// TIA Portal V20 export
// export: Created 2026-10-12T16:46:21.2512709Z, ExportSetting WithDefaults, DisplayName Totally Integrated Automation Portal, DisplayVersion V20 Update 6, DisplayName TIA Portal Openness, DisplayVersion V20 Update 6, DisplayName TIA Portal Version Control Interface, DisplayVersion V20 Update 6, DisplayName SINAMICS Startdrive Advanced, DisplayVersion V20 SP1 Update 2, DisplayName SINAMICS Startdrive G110M, G120, G120C, G120D, G120P, G115D, DisplayVersion V20 SP1 Update 2, DisplayName SINAMICS Startdrive G130, G150, S120, S150, SINAMICS MV, G220, S200, S210, DisplayVersion V20 SP1 Update 2, DisplayName STEP 7 Professional, DisplayVersion V20 Update 6, DisplayName STEP 7 Safety, DisplayVersion V20 Update 2, DisplayName WinCC Basic/Comfort/Advanced, DisplayVersion V20 Update 6, DisplayName WinCC Professional, DisplayVersion V20 Update 6, DisplayName WinCC Unified, DisplayVersion V20 Update 6
ORGANIZATION_BLOCK "Main"   // OB1, LAD, ProgramCycle
TITLE = "Main Program Sweep (Cycle)"
{ S7_Optimized_Access := 'TRUE' }
VERSION : 0.1
// stored: AutoNumber true, IsIECCheckEnabled false, SetENOAutomatically false
   VAR_INPUT
      Initial_Call : Bool;   // Initial call of this OB
      Remanence : Bool;   // =True, if remanent data are available
   END_VAR
   VAR_TEMP
      Lampentest_Ein : Bool;
      Blinktakt : Bool;
   END_VAR
BEGIN

REGION Network 1 (SCL): Eingaenge Lesen
   //KP8_1
   "FB_KP8_DB_1".KP8.Rohdaten.IB_Tasten := "KP8_1_IB_Tasten";
   "FB_KP8_DB_1".KP8.Rohdaten.IB_DI := "KP8_1_IB_DI";
   "FB_KP8_DB_1"();

   //KP8_2
   "FB_KP8_DB_2".KP8.Rohdaten.IB_Tasten := "KP8_2_IB_Tasten";
   "FB_KP8_DB_2".KP8.Rohdaten.IB_DI := "KP8_2_IB_DI";
   "FB_KP8_DB_2"();

   //KP8_3
   "FB_KP8_DB_3".KP8.Rohdaten.IB_Tasten := "KP8_3_IB_Tasten";
   "FB_KP8_DB_3".KP8.Rohdaten.IB_DI := "KP8_3_IB_DI";
   "FB_KP8_DB_3"();

   //KP8_4
   "FB_KP8_DB_4".KP8.Rohdaten.IB_Tasten := "KP8_4_IB_Tasten";
   "FB_KP8_DB_4".KP8.Rohdaten.IB_DI := "KP8_4_IB_DI";
   "FB_KP8_DB_4"();

   //KP8_5
   "FB_KP8_DB_5".KP8.Rohdaten.IB_Tasten := "KP8_5_IB_Tasten";
   "FB_KP8_DB_5".KP8.Rohdaten.IB_DI := "KP8_5_IB_DI";
   "FB_KP8_DB_5"();

   //KP8_6
   "FB_KP8_DB_6".KP8.Rohdaten.IB_Tasten := "KP8_6_IB_Tasten";
   "FB_KP8_DB_6".KP8.Rohdaten.IB_DI := "KP8_6_IB_DI";
   "FB_KP8_DB_6"();

   //KP8_7
   "FB_KP8_DB_7".KP8.Rohdaten.IB_Tasten := "KP8_7_IB_Tasten";
   "FB_KP8_DB_7".KP8.Rohdaten.IB_DI := "KP8_7_IB_DI";
   "FB_KP8_DB_7"();

   //KP8_8
   "FB_KP8_DB_8".KP8.Rohdaten.IB_Tasten := "KP8_8_IB_Tasten";
   "FB_KP8_DB_8".KP8.Rohdaten.IB_DI := "KP8_8_IB_DI";
   "FB_KP8_DB_8"();

   //KP8_9
   "FB_KP8_DB_9".KP8.Rohdaten.IB_Tasten := "KP8_9_IB_Tasten";
   "FB_KP8_DB_9".KP8.Rohdaten.IB_DI := "KP8_9_IB_DI";
   "FB_KP8_DB_9"();

   //KP8_10
   "FB_KP8_DB_10".KP8.Rohdaten.IB_Tasten := "KP8_10_IB_Tasten";
   "FB_KP8_DB_10".KP8.Rohdaten.IB_DI := "KP8_10_IB_DI";
   "FB_KP8_DB_10"();

   //KP8_11
   "FB_KP8_DB_11".KP8.Rohdaten.IB_Tasten := "KP8_11_IB_Tasten";
   "FB_KP8_DB_11".KP8.Rohdaten.IB_DI := "KP8_11_IB_DI";
   "FB_KP8_DB_11"();

   //KP8_12
   "FB_KP8_DB_12".KP8.Rohdaten.IB_Tasten := "KP8_12_IB_Tasten";
   "FB_KP8_DB_12".KP8.Rohdaten.IB_DI := "KP8_12_IB_DI";
   "FB_KP8_DB_12"();

   //KP8_13
   "FB_KP8_DB_13".KP8.Rohdaten.IB_Tasten := "KP8_13_IB_Tasten";
   "FB_KP8_DB_13".KP8.Rohdaten.IB_DI := "KP8_13_IB_DI";
   "FB_KP8_DB_13"();

   //KP8_14
   "FB_KP8_DB_14".KP8.Rohdaten.IB_Tasten := "KP8_14_IB_Tasten";
   "FB_KP8_DB_14".KP8.Rohdaten.IB_DI := "KP8_14_IB_DI";
   "FB_KP8_DB_14"();

   //KP8_15
   "FB_KP8_DB_15".KP8.Rohdaten.IB_Tasten := "KP8_15_IB_Tasten";
   "FB_KP8_DB_15".KP8.Rohdaten.IB_DI := "KP8_15_IB_DI";
   "FB_KP8_DB_15"();

   //KP8_16
   "FB_KP8_DB_16".KP8.Rohdaten.IB_Tasten := "KP8_16_IB_Tasten";
   "FB_KP8_DB_16".KP8.Rohdaten.IB_DI := "KP8_16_IB_DI";
   "FB_KP8_DB_16"();

   //KP8_17
   "FB_KP8_DB_17".KP8.Rohdaten.IB_Tasten := "KP8_17_IB_Tasten";
   "FB_KP8_DB_17".KP8.Rohdaten.IB_DI := "KP8_17_IB_DI";
   "FB_KP8_DB_17"();

   //KP8_18
   "FB_KP8_DB_18".KP8.Rohdaten.IB_Tasten := "KP8_18_IB_Tasten";
   "FB_KP8_DB_18".KP8.Rohdaten.IB_DI := "KP8_18_IB_DI";
   "FB_KP8_DB_18"();

   //KP8_19
   "FB_KP8_DB_19".KP8.Rohdaten.IB_Tasten := "KP8_19_IB_Tasten";
   "FB_KP8_DB_19".KP8.Rohdaten.IB_DI := "KP8_19_IB_DI";
   "FB_KP8_DB_19"();

   //KP8_20
   "FB_KP8_DB_20".KP8.Rohdaten.IB_Tasten := "KP8_20_IB_Tasten";
   "FB_KP8_DB_20".KP8.Rohdaten.IB_DI := "KP8_20_IB_DI";
   "FB_KP8_DB_20"();

   //KP8_21
   "FB_KP8_DB_21".KP8.Rohdaten.IB_Tasten := "KP8_21_IB_Tasten";
   "FB_KP8_DB_21".KP8.Rohdaten.IB_DI := "KP8_21_IB_DI";
   "FB_KP8_DB_21"();

   //KP8_22
   "FB_KP8_DB_22".KP8.Rohdaten.IB_Tasten := "KP8_22_IB_Tasten";
   "FB_KP8_DB_22".KP8.Rohdaten.IB_DI := "KP8_22_IB_DI";
   "FB_KP8_DB_22"();

   //KP8_23
   "FB_KP8_DB_23".KP8.Rohdaten.IB_Tasten := "KP8_23_IB_Tasten";
   "FB_KP8_DB_23".KP8.Rohdaten.IB_DI := "KP8_23_IB_DI";
   "FB_KP8_DB_23"();

   //KP8_24
   "FB_KP8_DB_24".KP8.Rohdaten.IB_Tasten := "KP8_24_IB_Tasten";
   "FB_KP8_DB_24".KP8.Rohdaten.IB_DI := "KP8_24_IB_DI";
   "FB_KP8_DB_24"();

   //KP8_25
   "FB_KP8_DB_25".KP8.Rohdaten.IB_Tasten := "KP8_25_IB_Tasten";
   "FB_KP8_DB_25".KP8.Rohdaten.IB_DI := "KP8_25_IB_DI";
   "FB_KP8_DB_25"();

   //KP8_26
   "FB_KP8_DB_26".KP8.Rohdaten.IB_Tasten := "KP8_26_IB_Tasten";
   "FB_KP8_DB_26".KP8.Rohdaten.IB_DI := "KP8_26_IB_DI";
   "FB_KP8_DB_26"();

   //KP8_27
   "FB_KP8_DB_27".KP8.Rohdaten.IB_Tasten := "KP8_27_IB_Tasten";
   "FB_KP8_DB_27".KP8.Rohdaten.IB_DI := "KP8_27_IB_DI";
   "FB_KP8_DB_27"();

   //KP8_28
   "FB_KP8_DB_28".KP8.Rohdaten.IB_Tasten := "KP8_28_IB_Tasten";
   "FB_KP8_DB_28".KP8.Rohdaten.IB_DI := "KP8_28_IB_DI";
   "FB_KP8_DB_28"();
END_REGION

REGION Network 2 (SCL): Badlogik
   "FB_Anlagensteuerung_DB"(Blink_Takt:="Clock_1Hz",
                            Clock_10Hz:="Clock_10Hz",
                            Not_Halt_Aktiv:=NOT "Not-Aus ist OK");
END_REGION

REGION Network 3 (SCL): Flexkraft
   // ----- 1) Eingänge aus Peripherie in den DB kopieren -----

   // FK_1 (IB500..IB531)
   "DB_FlexKraft_Data".FK_1.In.Reserved0            := "Flexkraft_1";    //IW500
   "DB_FlexKraft_Data".FK_1.In.StatusRegister       := "Flexkraft_2";    //IW502
   "DB_FlexKraft_Data".FK_1.In.WarningsRegister     := "Flexkraft_3";    //IW504
   "DB_FlexKraft_Data".FK_1.In.AlarmsRegister       := "Flexkraft_4";    //IW506
   "DB_FlexKraft_Data".FK_1.In.OutputVoltage        := "Flexkraft_5";    //IW508
   "DB_FlexKraft_Data".FK_1.In.OutputCurrent        := "Flexkraft_6";    //IW510
   "DB_FlexKraft_Data".FK_1.In.ProcessTime_HW       := "Flexkraft_7";    //IW512
   "DB_FlexKraft_Data".FK_1.In.ProcessTime_LW       := "Flexkraft_8";    //IW514
   "DB_FlexKraft_Data".FK_1.In.Ah_HW                := "Flexkraft_9";    //IW516
   "DB_FlexKraft_Data".FK_1.In.Ah_LW                := "Flexkraft_10";   //IW518

   // FK_2 (IB532..IB563)
   "DB_FlexKraft_Data".FK_2.In.Reserved0           := "Flexkraft_20";    //IW532
   "DB_FlexKraft_Data".FK_2.In.StatusRegister      := "Flexkraft_21";    //IW534
   "DB_FlexKraft_Data".FK_2.In.WarningsRegister    := "Flexkraft_22";    //IW536
   "DB_FlexKraft_Data".FK_2.In.AlarmsRegister      := "Flexkraft_23";    //IW538
   "DB_FlexKraft_Data".FK_2.In.OutputVoltage       := "Flexkraft_24";    //IW540
   "DB_FlexKraft_Data".FK_2.In.OutputCurrent       := "Flexkraft_25";    //IW542
   "DB_FlexKraft_Data".FK_2.In.ProcessTime_HW      := "Flexkraft_26";    //IW544
   "DB_FlexKraft_Data".FK_2.In.ProcessTime_LW      := "Flexkraft_27";    //IW546
   "DB_FlexKraft_Data".FK_2.In.Ah_HW               := "Flexkraft_28";    //IW548
   "DB_FlexKraft_Data".FK_2.In.Ah_LW               := "Flexkraft_29";    //IW550

   // FK_3 (IB564..IB595)
   "DB_FlexKraft_Data".FK_3.In.Reserved0           := "Flexkraft_30";    //IW564
   "DB_FlexKraft_Data".FK_3.In.StatusRegister      := "Flexkraft_31";    //IW566
   "DB_FlexKraft_Data".FK_3.In.WarningsRegister    := "Flexkraft_32";    //IW568
   "DB_FlexKraft_Data".FK_3.In.AlarmsRegister      := "Flexkraft_33";    //IW570
   "DB_FlexKraft_Data".FK_3.In.OutputVoltage       := "Flexkraft_34";    //IW572
   "DB_FlexKraft_Data".FK_3.In.OutputCurrent       := "Flexkraft_35";    //IW574
   "DB_FlexKraft_Data".FK_3.In.ProcessTime_HW      := "Flexkraft_36";    //IW576
   "DB_FlexKraft_Data".FK_3.In.ProcessTime_LW      := "Flexkraft_37";    //IW578
   "DB_FlexKraft_Data".FK_3.In.Ah_HW               := "Flexkraft_38";    //IW580
   "DB_FlexKraft_Data".FK_3.In.Ah_LW               := "Flexkraft_39";    //IW582

   // ----- 2) FB-Aufruf (1 Instanz pro Gerät) -----
   "FB_FlexKraft_DB"(bOn:="DB_Bad_Konfig".Bad_Konfig[40].GR_Aktiv,
                     bStartA:="DB_Bad_Konfig".Bad_Konfig[40].GR_Aktiv,
                     iSetVoltage_cV:="DB_Bad_Konfig".Bad_Konfig[40].GR_Spannung_Soll * 100,
                     iSetCurrent_raw:="DB_Bad_Konfig".Bad_Konfig[40].GR_Strom_Soll,
                     stDev:="DB_FlexKraft_Data".FK_1);

   "FB_FlexKraft_DB_1"(bOn:="DB_Bad_Konfig".Bad_Konfig[36].GR_Aktiv,
                       bStartA:="DB_Bad_Konfig".Bad_Konfig[36].GR_Aktiv,
                       iSetVoltage_cV:="DB_Bad_Konfig".Bad_Konfig[36].GR_Spannung_Soll * 100,
                       iSetCurrent_raw:="DB_Bad_Konfig".Bad_Konfig[36].GR_Strom_Soll,
                       stDev:="DB_FlexKraft_Data".FK_2);

   "FB_FlexKraft_DB_2"(bOn:="DB_Bad_Konfig".Bad_Konfig[31].GR_Aktiv,
                       bStartA:="DB_Bad_Konfig".Bad_Konfig[31].GR_Aktiv,
                       iSetVoltage_cV:="DB_Bad_Konfig".Bad_Konfig[31].GR_Spannung_Soll * 100,
                       iSetCurrent_raw:="DB_Bad_Konfig".Bad_Konfig[31].GR_Strom_Soll,
                       stDev:="DB_FlexKraft_Data".FK_3);


   // ----- 3) Ausgänge aus dem DB in die Peripherie kopieren -----

   // FK_1 (QB500..QB531)
   "Flexkraft_11"    := "DB_FlexKraft_Data".FK_1.Out.PageNo;                 //QW500
   "Flexkraft_12"    := "DB_FlexKraft_Data".FK_1.Out.ControlRegister;        //QW502
   "Flexkraft_13"    := "DB_FlexKraft_Data".FK_1.Out.SetVoltage;             //QW504
   "Flexkraft_14"    := "DB_FlexKraft_Data".FK_1.Out.SetCurrent;             //QW506
   "Flexkraft_15"    := "DB_FlexKraft_Data".FK_1.Out.ProcessTimerLimit_HW;   //QW508
   "Flexkraft_16"    := "DB_FlexKraft_Data".FK_1.Out.ProcessTimerLimit_LW;   //QW510
   "Flexkraft_17"    := "DB_FlexKraft_Data".FK_1.Out.AhLimit_HW;             //QW512
   "Flexkraft_18"    := "DB_FlexKraft_Data".FK_1.Out.AhLimit_LW;             //QW514
   "Flexkraft_19"    := "DB_FlexKraft_Data".FK_1.Out.Startramp;              //QW516

   // FK_2 (QB532..QB563)
   "Flexkraft_40"    :="DB_FlexKraft_Data".FK_2.Out.PageNo;                  //QW532
   "Flexkraft_41"    :="DB_FlexKraft_Data".FK_2.Out.ControlRegister;         //QW534
   "Flexkraft_42"    :="DB_FlexKraft_Data".FK_2.Out.SetVoltage;              //QW536
   "Flexkraft_43"    :="DB_FlexKraft_Data".FK_2.Out.SetCurrent;              //QW538
   "Flexkraft_44"    :="DB_FlexKraft_Data".FK_2.Out.ProcessTimerLimit_HW;    //QW540
   "Flexkraft_45"    :="DB_FlexKraft_Data".FK_2.Out.ProcessTimerLimit_LW;    //QW542
   "Flexkraft_46"    :="DB_FlexKraft_Data".FK_2.Out.AhLimit_HW;              //QW544
   "Flexkraft_49"    :="DB_FlexKraft_Data".FK_2.Out.AhLimit_LW;              //QW546
   "Flexkraft_48"    :="DB_FlexKraft_Data".FK_2.Out.Startramp;               //QW548

   // FK_3 (QB564..QB595)
   "Flexkraft_47"    :="DB_FlexKraft_Data".FK_3.Out.PageNo;                  //QW564
   "Flexkraft_50"    :="DB_FlexKraft_Data".FK_3.Out.ControlRegister;         //QW566
   "Flexkraft_51"    :="DB_FlexKraft_Data".FK_3.Out.SetVoltage;              //QW568
   "Flexkraft_52"    :="DB_FlexKraft_Data".FK_3.Out.SetCurrent;              //QW570
   "Flexkraft_54"    :="DB_FlexKraft_Data".FK_3.Out.ProcessTimerLimit_HW;    //QW572
   "Flexkraft_53"    :="DB_FlexKraft_Data".FK_3.Out.ProcessTimerLimit_LW;    //QW574
   "Flexkraft_55"    :="DB_FlexKraft_Data".FK_3.Out.AhLimit_HW;              //QW576
   "Flexkraft_56"    :="DB_FlexKraft_Data".FK_3.Out.AhLimit_LW;              //QW578
   "Flexkraft_57"    :="DB_FlexKraft_Data".FK_3.Out.Startramp;               //QW580
END_REGION

REGION Network 4 (SCL): Ausgaenge schreiben

   //KP8_1
   "FB_KP8_DB_1"();
   "KP8_1_QB_Rot" := "FB_KP8_DB_1".KP8.Rohdaten.QB_Rot;
   "KP8_1_QB_Gruen" := "FB_KP8_DB_1".KP8.Rohdaten.QB_Gruen;
   "KP8_1_QB_Blau" := "FB_KP8_DB_1".KP8.Rohdaten.QB_Blau;
   "KP8_1_QB_DO" := "FB_KP8_DB_1".KP8.Rohdaten.QB_DO;

   //KP8_2
   "FB_KP8_DB_2"();
   "KP8_2_QB_Rot" := "FB_KP8_DB_2".KP8.Rohdaten.QB_Rot;
   "KP8_2_QB_Gruen" := "FB_KP8_DB_2".KP8.Rohdaten.QB_Gruen;
   "KP8_2_QB_Blau" := "FB_KP8_DB_2".KP8.Rohdaten.QB_Blau;
   "KP8_2_QB_DO" := "FB_KP8_DB_2".KP8.Rohdaten.QB_DO;

   //KP8_3
   "FB_KP8_DB_3"();
   "KP8_3_QB_Rot" := "FB_KP8_DB_3".KP8.Rohdaten.QB_Rot;
   "KP8_3_QB_Gruen" := "FB_KP8_DB_3".KP8.Rohdaten.QB_Gruen;
   "KP8_3_QB_Blau" := "FB_KP8_DB_3".KP8.Rohdaten.QB_Blau;
   "KP8_3_QB_DO" := "FB_KP8_DB_3".KP8.Rohdaten.QB_DO;

   //KP8_4
   "FB_KP8_DB_4"();
   "KP8_4_QB_Rot" := "FB_KP8_DB_4".KP8.Rohdaten.QB_Rot;
   "KP8_4_QB_Gruen" := "FB_KP8_DB_4".KP8.Rohdaten.QB_Gruen;
   "KP8_4_QB_Blau" := "FB_KP8_DB_4".KP8.Rohdaten.QB_Blau;
   "KP8_4_QB_DO" := "FB_KP8_DB_4".KP8.Rohdaten.QB_DO;

   //KP8_5
   "FB_KP8_DB_5"();
   "KP8_5_QB_Rot" := "FB_KP8_DB_5".KP8.Rohdaten.QB_Rot;
   "KP8_5_QB_Gruen" := "FB_KP8_DB_5".KP8.Rohdaten.QB_Gruen;
   "KP8_5_QB_Blau" := "FB_KP8_DB_5".KP8.Rohdaten.QB_Blau;
   "KP8_5_QB_DO" := "FB_KP8_DB_5".KP8.Rohdaten.QB_DO;

   //KP8_6
   "FB_KP8_DB_6"();
   "KP8_6_QB_Rot" := "FB_KP8_DB_6".KP8.Rohdaten.QB_Rot;
   "KP8_6_QB_Gruen" := "FB_KP8_DB_6".KP8.Rohdaten.QB_Gruen;
   "KP8_6_QB_Blau" := "FB_KP8_DB_6".KP8.Rohdaten.QB_Blau;
   "KP8_6_QB_DO" := "FB_KP8_DB_6".KP8.Rohdaten.QB_DO;

   //KP8_7
   "FB_KP8_DB_7"();
   "KP8_7_QB_Rot" := "FB_KP8_DB_7".KP8.Rohdaten.QB_Rot;
   "KP8_7_QB_Gruen" := "FB_KP8_DB_7".KP8.Rohdaten.QB_Gruen;
   "KP8_7_QB_Blau" := "FB_KP8_DB_7".KP8.Rohdaten.QB_Blau;
   "KP8_7_QB_DO" := "FB_KP8_DB_7".KP8.Rohdaten.QB_DO;

   //KP8_8
   "FB_KP8_DB_8"();
   "KP8_8_QB_Rot" := "FB_KP8_DB_8".KP8.Rohdaten.QB_Rot;
   "KP8_8_QB_Gruen" := "FB_KP8_DB_8".KP8.Rohdaten.QB_Gruen;
   "KP8_8_QB_Blau" := "FB_KP8_DB_8".KP8.Rohdaten.QB_Blau;
   "KP8_8_QB_DO" := "FB_KP8_DB_8".KP8.Rohdaten.QB_DO;

   //KP8_9
   "FB_KP8_DB_9"();
   "KP8_9_QB_Rot" := "FB_KP8_DB_9".KP8.Rohdaten.QB_Rot;
   "KP8_9_QB_Gruen" := "FB_KP8_DB_9".KP8.Rohdaten.QB_Gruen;
   "KP8_9_QB_Blau" := "FB_KP8_DB_9".KP8.Rohdaten.QB_Blau;
   "KP8_9_QB_DO" := "FB_KP8_DB_9".KP8.Rohdaten.QB_DO;

   //KP8_10
   "FB_KP8_DB_10"();
   "KP8_10_QB_Rot" := "FB_KP8_DB_10".KP8.Rohdaten.QB_Rot;
   "KP8_10_QB_Gruen" := "FB_KP8_DB_10".KP8.Rohdaten.QB_Gruen;
   "KP8_10_QB_Blau" := "FB_KP8_DB_10".KP8.Rohdaten.QB_Blau;
   "KP8_10_QB_DO" := "FB_KP8_DB_10".KP8.Rohdaten.QB_DO;

   //KP8_11
   "FB_KP8_DB_11"();
   "KP8_11_QB_Rot" := "FB_KP8_DB_11".KP8.Rohdaten.QB_Rot;
   "KP8_11_QB_Gruen" := "FB_KP8_DB_11".KP8.Rohdaten.QB_Gruen;
   "KP8_11_QB_Blau" := "FB_KP8_DB_11".KP8.Rohdaten.QB_Blau;
   "KP8_11_QB_DO" := "FB_KP8_DB_11".KP8.Rohdaten.QB_DO;

   //KP8_12
   "FB_KP8_DB_12"();
   "KP8_12_QB_Rot" := "FB_KP8_DB_12".KP8.Rohdaten.QB_Rot;
   "KP8_12_QB_Gruen" := "FB_KP8_DB_12".KP8.Rohdaten.QB_Gruen;
   "KP8_12_QB_Blau" := "FB_KP8_DB_12".KP8.Rohdaten.QB_Blau;
   "KP8_12_QB_DO" := "FB_KP8_DB_12".KP8.Rohdaten.QB_DO;

   //KP8_13
   "FB_KP8_DB_13"();
   "KP8_13_QB_Rot" := "FB_KP8_DB_13".KP8.Rohdaten.QB_Rot;
   "KP8_13_QB_Gruen" := "FB_KP8_DB_13".KP8.Rohdaten.QB_Gruen;
   "KP8_13_QB_Blau" := "FB_KP8_DB_13".KP8.Rohdaten.QB_Blau;
   "KP8_13_QB_DO" := "FB_KP8_DB_13".KP8.Rohdaten.QB_DO;

   //KP8_14
   "FB_KP8_DB_14"();
   "KP8_14_QB_Rot" := "FB_KP8_DB_14".KP8.Rohdaten.QB_Rot;
   "KP8_14_QB_Gruen" := "FB_KP8_DB_14".KP8.Rohdaten.QB_Gruen;
   "KP8_14_QB_Blau" := "FB_KP8_DB_14".KP8.Rohdaten.QB_Blau;
   "KP8_14_QB_DO" := "FB_KP8_DB_14".KP8.Rohdaten.QB_DO;

   //KP8_15
   "FB_KP8_DB_15"();
   "KP8_15_QB_Rot" := "FB_KP8_DB_15".KP8.Rohdaten.QB_Rot;
   "KP8_15_QB_Gruen" := "FB_KP8_DB_15".KP8.Rohdaten.QB_Gruen;
   "KP8_15_QB_Blau" := "FB_KP8_DB_15".KP8.Rohdaten.QB_Blau;
   "KP8_15_QB_DO" := "FB_KP8_DB_15".KP8.Rohdaten.QB_DO;

   //KP8_16
   "FB_KP8_DB_16"();
   "KP8_16_QB_Rot" := "FB_KP8_DB_16".KP8.Rohdaten.QB_Rot;
   "KP8_16_QB_Gruen" := "FB_KP8_DB_16".KP8.Rohdaten.QB_Gruen;
   "KP8_16_QB_Blau" := "FB_KP8_DB_16".KP8.Rohdaten.QB_Blau;
   "KP8_16_QB_DO" := "FB_KP8_DB_16".KP8.Rohdaten.QB_DO;

   //KP8_17
   "FB_KP8_DB_17"();
   "KP8_17_QB_Rot" := "FB_KP8_DB_17".KP8.Rohdaten.QB_Rot;
   "KP8_17_QB_Gruen" := "FB_KP8_DB_17".KP8.Rohdaten.QB_Gruen;
   "KP8_17_QB_Blau" := "FB_KP8_DB_17".KP8.Rohdaten.QB_Blau;
   "KP8_17_QB_DO" := "FB_KP8_DB_17".KP8.Rohdaten.QB_DO;

   //KP8_18
   "FB_KP8_DB_18"();
   "KP8_18_QB_Rot" := "FB_KP8_DB_18".KP8.Rohdaten.QB_Rot;
   "KP8_18_QB_Gruen" := "FB_KP8_DB_18".KP8.Rohdaten.QB_Gruen;
   "KP8_18_QB_Blau" := "FB_KP8_DB_18".KP8.Rohdaten.QB_Blau;
   "KP8_18_QB_DO" := "FB_KP8_DB_18".KP8.Rohdaten.QB_DO;

   //KP8_19
   "FB_KP8_DB_19"();
   "KP8_19_QB_Rot" := "FB_KP8_DB_19".KP8.Rohdaten.QB_Rot;
   "KP8_19_QB_Gruen" := "FB_KP8_DB_19".KP8.Rohdaten.QB_Gruen;
   "KP8_19_QB_Blau" := "FB_KP8_DB_19".KP8.Rohdaten.QB_Blau;
   "KP8_19_QB_DO" := "FB_KP8_DB_19".KP8.Rohdaten.QB_DO;

   //KP8_20
   "FB_KP8_DB_20"();
   "KP8_20_QB_Rot" := "FB_KP8_DB_20".KP8.Rohdaten.QB_Rot;
   "KP8_20_QB_Gruen" := "FB_KP8_DB_20".KP8.Rohdaten.QB_Gruen;
   "KP8_20_QB_Blau" := "FB_KP8_DB_20".KP8.Rohdaten.QB_Blau;
   "KP8_20_QB_DO" := "FB_KP8_DB_20".KP8.Rohdaten.QB_DO;

   //KP8_21
   "FB_KP8_DB_21"();
   "KP8_21_QB_Rot" := "FB_KP8_DB_21".KP8.Rohdaten.QB_Rot;
   "KP8_21_QB_Gruen" := "FB_KP8_DB_21".KP8.Rohdaten.QB_Gruen;
   "KP8_21_QB_Blau" := "FB_KP8_DB_21".KP8.Rohdaten.QB_Blau;
   "KP8_21_QB_DO" := "FB_KP8_DB_21".KP8.Rohdaten.QB_DO;

   //KP8_22
   "FB_KP8_DB_22"();
   "KP8_22_QB_Rot" := "FB_KP8_DB_22".KP8.Rohdaten.QB_Rot;
   "KP8_22_QB_Gruen" := "FB_KP8_DB_22".KP8.Rohdaten.QB_Gruen;
   "KP8_22_QB_Blau" := "FB_KP8_DB_22".KP8.Rohdaten.QB_Blau;
   "KP8_22_QB_DO" := "FB_KP8_DB_22".KP8.Rohdaten.QB_DO;

   //KP8_23
   "FB_KP8_DB_23"();
   "KP8_23_QB_Rot" := "FB_KP8_DB_23".KP8.Rohdaten.QB_Rot;
   "KP8_23_QB_Gruen" := "FB_KP8_DB_23".KP8.Rohdaten.QB_Gruen;
   "KP8_23_QB_Blau" := "FB_KP8_DB_23".KP8.Rohdaten.QB_Blau;
   "KP8_23_QB_DO" := "FB_KP8_DB_23".KP8.Rohdaten.QB_DO;

   //KP8_24
   "FB_KP8_DB_24"();
   "KP8_24_QB_Rot" := "FB_KP8_DB_24".KP8.Rohdaten.QB_Rot;
   "KP8_24_QB_Gruen" := "FB_KP8_DB_24".KP8.Rohdaten.QB_Gruen;
   "KP8_24_QB_Blau" := "FB_KP8_DB_24".KP8.Rohdaten.QB_Blau;
   "KP8_24_QB_DO" := "FB_KP8_DB_24".KP8.Rohdaten.QB_DO;

   //KP8_25
   "FB_KP8_DB_25"();
   "KP8_25_QB_Rot" := "FB_KP8_DB_25".KP8.Rohdaten.QB_Rot;
   "KP8_25_QB_Gruen" := "FB_KP8_DB_25".KP8.Rohdaten.QB_Gruen;
   "KP8_25_QB_Blau" := "FB_KP8_DB_25".KP8.Rohdaten.QB_Blau;
   "KP8_25_QB_DO" := "FB_KP8_DB_25".KP8.Rohdaten.QB_DO;

   //KP8_26
   "FB_KP8_DB_26"();
   "KP8_26_QB_Rot" := "FB_KP8_DB_26".KP8.Rohdaten.QB_Rot;
   "KP8_26_QB_Gruen" := "FB_KP8_DB_26".KP8.Rohdaten.QB_Gruen;
   "KP8_26_QB_Blau" := "FB_KP8_DB_26".KP8.Rohdaten.QB_Blau;
   "KP8_26_QB_DO" := "FB_KP8_DB_26".KP8.Rohdaten.QB_DO;

   //KP8_27
   "FB_KP8_DB_27"();
   "KP8_27_QB_Rot" := "FB_KP8_DB_27".KP8.Rohdaten.QB_Rot;
   "KP8_27_QB_Gruen" := "FB_KP8_DB_27".KP8.Rohdaten.QB_Gruen;
   "KP8_27_QB_Blau" := "FB_KP8_DB_27".KP8.Rohdaten.QB_Blau;
   "KP8_27_QB_DO" := "FB_KP8_DB_27".KP8.Rohdaten.QB_DO;

   //KP8_28
   "FB_KP8_DB_28"();
   "KP8_28_QB_Rot" := "FB_KP8_DB_28".KP8.Rohdaten.QB_Rot;
   "KP8_28_QB_Gruen" := "FB_KP8_DB_28".KP8.Rohdaten.QB_Gruen;
   "KP8_28_QB_Blau" := "FB_KP8_DB_28".KP8.Rohdaten.QB_Blau;
   "KP8_28_QB_DO" := "FB_KP8_DB_28".KP8.Rohdaten.QB_DO;
END_REGION

REGION Network 5 (SCL): Fehlermeldungen
   "FC_Fehlermeldungen"();
END_REGION

REGION Network 6 (SCL): Not-Halt
   "FC_Not_Halt"(NOT "Not-Aus ist OK");
END_REGION

REGION Network 7 (SCL): Not-Aus Reset
       "Not-Aus Reset" := "DB_IPC_to_CPU".Not_Halt_Reset;     // %Q4.7
END_REGION
END_ORGANIZATION_BLOCK
